// TIA Portal V19 export
TYPE "ST_REER_INPUT_BYTE"
   STRUCT
      INPUT : Array[0..32] of Byte;
   END_STRUCT;
END_TYPE
